FUNCTION_BLOCK ProcessDataManager EXTENDS TcoData.TcoDataExchange
VAR
	//this variable has to called "_data" - PC app will access this variable by its name.
	 {attribute clr [Container(Layout.Tabs)]}
     {attribute clr [Group(Layout.Scroll)]}
	_data : Station001_ProductionData := (Parent := THIS^);
END_VAR

SUPER^();

//Set default values in case that no setting has been loaded into the PLC yet.
//IF _data.DimX.Mininum = 0 AND _data.DimX.Maximum = 0 THEN
//    _data.DimX.Mininum :=
//        0.95 * MAIN._app._station001._components._dimXsim.inMinValue + 0.05 * MAIN._app._station001._components._dimXsim.inMaxValue;

//    _data.DimX.Maximum :=
//        0.05 * MAIN._app._station001._components._dimXsim.inMinValue + 0.95 * MAIN._app._station001._components._dimXsim.inMaxValue;
//END_IF

//IF _data.DimY.Mininum = 0 AND _data.DimY.Maximum = 0 THEN
//    _data.DimY.Mininum :=
//        0.95 * MAIN._app._station001._components._dimYsim.inMinValue + 0.05 * MAIN._app._station001._components._dimYsim.inMaxValue;

//    _data.DimY.Maximum :=
//        0.05 * MAIN._app._station001._components._dimYsim.inMinValue + 0.95 * MAIN._app._station001._components._dimYsim.inMaxValue;
//END_IF

//IF _data.DimZ.Mininum = 0 AND _data.DimZ.Maximum = 0 THEN
//    _data.DimZ.Mininum :=
//        0.95 * MAIN._app._station001._components._dimZsim.inMinValue + 0.05 * MAIN._app._station001._components._dimZsim.inMaxValue;

//    _data.DimZ.Maximum :=
//        0.05 * MAIN._app._station001._components._dimZsim.inMinValue + 0.95 * MAIN._app._station001._components._dimZsim.inMaxValue;
//END_IF

METHOD SetDataResult
VAR_INPUT
	Result : TcoComprehensiveResult;
END_VAR
_data.Result := Result;
END_METHOD

METHOD SetRecipe
VAR_INPUT
	RecipeName:STRING;
END_VAR
_data.RecipeName := RecipeName;
END_METHOD

END_FUNCTION_BLOCK

(* stored: Version 1.1.0.1, ProductVersion 3.1.4024.9
   POU ProcessDataManager: Id {ef58d043-6bbe-480b-9350-92a4de31085d}, SpecialFunc None
   Method SetDataResult: Id {18eeae59-e657-0c7b-3528-07fbaa61af6f}
   Method SetRecipe: Id {311d426e-c67b-0715-0737-1237a18f8640} *)
